TYPE "ST_TimeQuality"
VERSION : 0.1
   STRUCT
      "Available" : Bool;
      "Synchronized" : Bool;
      "Source" : String[32];
      "OffsetUs" : DInt;
      "LastSyncAt" : LDT;
      "ObservedAt" : LDT;
   END_STRUCT;
END_TYPE
